Universal Robots URScript: Pick1.script

def Pick1():
  # Global parameters:
  global speed_ms    = 0.250
  global speed_rads  = 0.750
  global accel_mss   = 1.200
  global accel_radss = 1.200
  global blend_radius_m = 0.001
  global ref_frame = p[0,0,0,0,0,0]

  #
  # TO REMOVE HEADER:
  # Go to "Program" -> "Post-Processor Editor"
  # Select "Universal Robots"
  # Set "INCLUDE_HEADER" to "False"
  #
  #--------------------------
  # Add any default subprograms here
  # For example, to drive a gripper as a program call:
  # def Gripper_Open():
  #   ...
  # end
  #
  # Example to drive a spray gun:
  def SprayOn(value):
    # use the value as an output:
    DO_SPRAY = 5
    if value == 0:
      set_standard_digital_out(DO_SPRAY, False)
    else:
      set_standard_digital_out(DO_SPRAY, True)
    end
  end

  # Example to drive an extruder:
  def Extruder(value):
    # use the value as an output:
    if value < 0:
      # stop extruder
    else:
      # start extruder
    end
  end

  # Example to move an external axis
  def MoveAxis(value):
    # use the value as an output:
    DO_AXIS_1 = 1
    DI_AXIS_1 = 1
    if value <= 0:
      set_standard_digital_out(DO_AXIS_1, False)

      # Wait for digital input to change state
      #while (get_standard_digital_in(DI_AXIS_1) != False):
      #  sync()
      #end
    else:
      set_standard_digital_out(DO_AXIS_1, True)

      # Wait for digital input to change state
      #while (get_standard_digital_in(DI_AXIS_1) != True):
      #  sync()
      #end
    end
  end
  #--------------------------

  # Subprogram Gripper1PickInput
  def Gripper1PickInput():
    CloseGripper1()
    # Attach to Gripper1
    # Attach to Gripper1
  end

  # Subprogram CloseGripper1
  def CloseGripper1():
    movej([0.698132, 0.000000, 0.000000, 0.000000, 0.000000, 0.000000],accel_radss,speed_rads,0,0.001)
  end


  # Main program:
  # Program generated by VerticalBot Studio for UR10e on 25/10/2026 12:00:00
  # Using nominal kinematics.
  ref_frame = p[-0.500000, -0.590000, 0.300000, 0.000000, 0.000000, 0.000000]
  set_tcp(p[0.145000, 0.000000, 0.130000, 0.613943, 0.613943, 1.482190])
  movej([-5.367551, -2.005139, 2.365131, -3.501602, -1.701036, -0.000000],accel_radss,speed_rads,0,0.001)
  movel(pose_trans(ref_frame,p[0.192500, 0.192500, 0.115000, -2.221441, -0.000000, 2.221441]),accel_mss,speed_ms,0,0) # end trace
  Gripper1PickInput()
  movel(pose_trans(ref_frame,p[0.192500, 0.192500, 0.355000, -2.221441, 0.000000, 2.221441]),accel_mss,speed_ms,0,0.001)
  # End of main program
end

Pick1()
